TYPE TwinSafeOut_PlcIn :
STRUCT
	FB_Err			: BOOL;
	COM_Err			: BOOL;
	OUT_Err			: BOOL;
	Other_Err		: BOOL;
	InRun			: BOOL;
	//ES_State		: BOOL;

END_STRUCT
END_TYPE

(* stored: Version 1.1.0.1, ProductVersion 3.1.4024.13
   DUT TwinSafeOut_PlcIn: Id {a5fc3abe-d301-4f8d-ae1b-61d2611fd80a} *)
